Fanuc KAREL source: KA00195.KL

PROGRAM KA00195
%NOLOCKGROUP
VAR
  SRC: ARRAY[4] OF SHORT
  DST: ARRAY[4] OF SHORT
BEGIN
  DST = SRC
END KA00195
